INTERFACE I_Actuator EXTENDS I_Diagnosable, I_Resettable

METHOD Extend
END_METHOD

METHOD Retract
END_METHOD

PROPERTY IsExtended : BOOL
GET
END_GET
END_PROPERTY

PROPERTY IsRetracted : BOOL
GET
END_GET
END_PROPERTY

END_INTERFACE

(* stored: Version 1.1.0.1
   Itf I_Actuator: Id {e5a864e7-19b8-4986-8afb-1fd2e859fd00}
   Method Extend: Id {b1118beb-73e5-4aff-8aed-2c76d9743b9d}
   Method Retract: Id {9d53b4e8-2d59-4539-8cef-807f7bbeb199}
   Property IsExtended: Id {16afcaa6-6f34-4f41-a661-c2fb890ab126}
   Get Get: Id {c93f0d5f-617d-4258-9682-e1538dbc1c96}
   Property IsRetracted: Id {905338a5-bd2a-48ec-929b-ee3cc87bc915}
   Get Get: Id {5c148518-0383-4853-a6c3-89c56b37f140} *)
